TYPE st_LineTargetValves :
STRUCT
	valTankA				:	E_Pis_Name	;
	valTankB				:	E_Pis_Name	;
	valDrain				:	E_Pis_Name	;
	valCIP					:	E_Pis_Name	;
	valTankA_Pipe			:	E_Pis_Name	;
	valTankB_Pipe			:	E_Pis_Name	;
END_STRUCT
END_TYPE

(* stored: Version 1.1.0.1, ProductVersion 3.1.4024.12
   DUT st_LineTargetValves: Id {2ad8f729-2c39-458f-901e-b914d6de7ecc} *)
